INTERFACE I_IoBase

METHOD Update
VAR_INPUT
END_VAR
END_METHOD

END_INTERFACE

(* stored: Version 1.1.0.1
   Itf I_IoBase: Id {a414fd6f-6217-4683-a2ae-eb3302fcd51a}
   Method Update: Id {1d304fa5-17b2-4307-9b2b-3b02dc801f3f} *)
